(* IEC 61131-3 sources: 2026_Projet_YGO_ExcavatriceDragage/CODE/SYSTEM, 3 files *)

(* ---- GVL_BUS.st ---- *)
(* ═══════════════════════════════════════════════════════════════
   🗑️ GVL_BUS — Obsolete / Archive
   ───────────────────────────────────────────────────────────────
   Note : Suite à la décision d'architecture D2, la surveillance par
   dégradation de bus (GVL_BusHealth / E_DegradationLevel) a été
   supprimée. Ce fichier est conservé uniquement pour archive de structure.
   ═══════════════════════════════════════════════════════════════ *)
VAR_GLOBAL
    // GVL obsolète - non référencé par PRG_MAIN
END_VAR

(* ---- GVL_Machine_Stub.st ---- *)
(* ═══════════════════════════════════════════════════════════════
   🏭 GVL_Machine_Stub — Variables IHM transverses machine (Lot A mise en service)
   ───────────────────────────────────────────────────────────────
   📄 Doc métier : DOC/AF_Partie3_Template_FB_Commun_v1.3.md §5 (bouton général)
   🎯 `MachineReset_IHM` : bouton acquittement GÉNÉRAL (front) — distribué à TOUTES les
      instances (diag, modes, safety, winch, chariot, winchsync + OR-é avec les boutons
      par codeur M1/M2_Reset_IHM). Partie3 §5 : « bouton général ».
   🔧 CORRECTIF (2026-07-03quindecies) : `PowerCutOffCmd` retiré — relais réel câblé en
      I/O Mapping (`PowerCutOff_RQ`), voir PRG_MAIN.st §8.
   🔴 TOUJOURS STUB (pas de vrai bouton IHM câblé) : `MachineReset_IHM` se force en vue
      instance CODESYS (TRUE puis FALSE = front).
   ═══════════════════════════════════════════════════════════════ *)

// === DECLARATION (à coller dans la partie déclaration du GVL GVL_Machine_Stub) ===

VAR_GLOBAL
    // 🔑 Acquittement général machine (front) — acquitte TOUS les FB d'un coup
    MachineReset_IHM : BOOL;   // 🖥️ À mapper bouton IHM — basculer TRUE puis FALSE pour simuler l'appui
END_VAR

(* ---- FB_CycleTime.st ---- *)
(* ═══════════════════════════════════════════════════════════════
   ⏱️ FB_CycleTime — Mesure du temps de cycle réel de la tâche
   ═══════════════════════════════════════════════════════════════ *)
FUNCTION_BLOCK FB_CycleTime
VAR_INPUT
    DefaultValueS : REAL := 0.004; (* Valeur de secours par défaut (ex. 4ms) *)
END_VAR
VAR_OUTPUT
    CycleTimeS    : REAL;          (* Temps écoulé réel calculé (secondes) *)
END_VAR
VAR
    TimeCurrent   : TIME;          (* Temps système actuel *)
    TimeLast      : TIME;          (* Empreinte de temps du cycle précédent *)
    DeltaTimeMs   : UDINT;         (* Écart brut calculé (ms) *)
    InitDone      : BOOL;          (* Drapeau d'initialisation du premier cycle *)
END_VAR

// 1. ACQUISITION DU TEMPS SYSTÈME
TimeCurrent := TIME();

// 2. INITIALISATION UNIQUE AU PREMIER CYCLE
IF NOT InitDone THEN
    TimeLast := TimeCurrent;
    InitDone := TRUE;
    CycleTimeS := DefaultValueS;
    RETURN;
END_IF;

// 3. CALCUL DU DELTA EN MILLISECONDES
DeltaTimeMs := TIME_TO_UDINT(TimeCurrent - TimeLast);

// 4. CONVERSION ET CHARGE DE SECOURS
IF DeltaTimeMs > 0 THEN
    CycleTimeS := UDINT_TO_REAL(DeltaTimeMs) / 1000.0;
ELSE
    CycleTimeS := DefaultValueS;
END_IF;

// 5. ARCHIVAGE POUR LE PROCHAIN CYCLE
TimeLast := TimeCurrent;
